PROGRAM main
  VAR
    B1 AT %IX0.0   : BOOL; (* sensor de cajas *)
    KM1 AT %QX0.0  : BOOL; (* banda (bobina 00001 para la PC) *)
    CAJAS AT %MW0  : INT; (* holding 40001: cajas contadas *)
    MARCHA AT %MW1 : INT; (* holding 40002: marcha, la escribe la PC *)
    META AT %MW2   : INT; (* holding 40003: meta de cajas, la escribe la PC *)
    F_CAJA         : R_TRIG;
    CAJA           : BOOL; (* flanco de B1 *)
  END_VAR
  VAR  (* added by the conversion: wires and edge detectors of the diagram *)
    _ADD7_OUT : INT;
    _SEL4_OUT : INT;
    _GT13_OUT : BOOL;
    _GE16_OUT : BOOL;
    _AND12_OUT : BOOL;
    _SEL11_OUT : INT;
    _NE22_OUT : BOOL;
  END_VAR

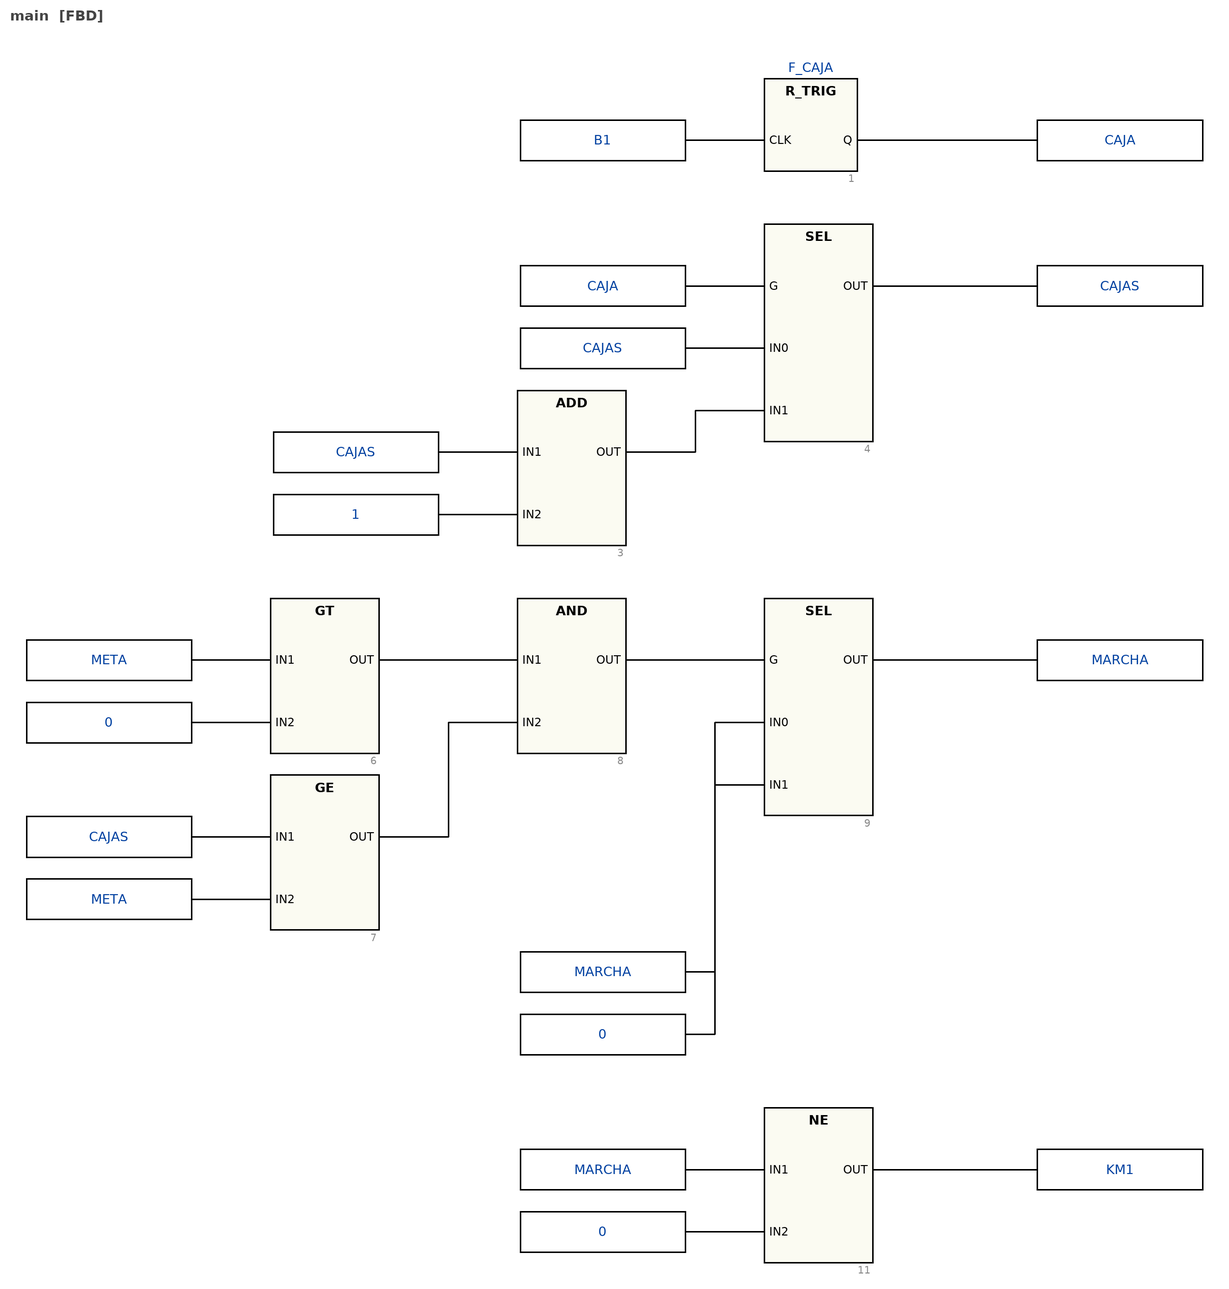
(* FBD diagram, written out as Structured Text *)
F_CAJA(CLK := B1);
CAJA := F_CAJA.Q;
_ADD7_OUT := CAJAS + 1;
_SEL4_OUT := SEL(CAJA, CAJAS, _ADD7_OUT);
CAJAS := _SEL4_OUT;
_GT13_OUT := META > 0;
_GE16_OUT := CAJAS >= META;
_AND12_OUT := _GT13_OUT AND _GE16_OUT;
_SEL11_OUT := SEL(_AND12_OUT, MARCHA, 0);
MARCHA := _SEL11_OUT;
_NE22_OUT := MARCHA <> 0;
KM1 := _NE22_OUT;
END_PROGRAM
